{attribute 'qualified_only'}
{attribute 'strict'}
TYPE E_Tank_Level :
(
	eEmpty := 0,
	eLL,
	eHL,
	eERROR
	
);
END_TYPE

(* stored: Version 1.1.0.1, ProductVersion 3.1.4024.12
   DUT E_Tank_Level: Id {e3fd1449-4f5d-487b-9760-17039c463210} *)
